// TIA Portal V20 export
// export: Created 2026-10-19T18:06:52.8062617Z, ExportSetting WithDefaults, DisplayName Totally Integrated Automation Portal, DisplayVersion V20 Update 6, DisplayName TIA Portal Openness, DisplayVersion V20 Update 6, DisplayName TIA Portal Version Control Interface, DisplayVersion V20 Update 6, DisplayName SINAMICS Startdrive Advanced, DisplayVersion V20 SP1, DisplayName SINAMICS Startdrive G130, G150, S120, S150, SINAMICS MV, G220, S200, S210, DisplayVersion V20 SP1, DisplayName SINAMICS Startdrive G110M, G120, G120C, G120D, G120P, G115D, DisplayVersion V20 SP1, DisplayName STEP 7 Professional, DisplayVersion V20 Update 6, DisplayName STEP 7 Safety, DisplayVersion V20 Update 2, DisplayName WinCC Basic/Comfort/Advanced, DisplayVersion V20 Update 6, DisplayName WinCC Unified, DisplayVersion V20 Update 6
DATA_BLOCK "SAI_IND_SpanAdjust_DB"   // DB113
VERSION : 0.1
// stored: AutoNumber true, DBAccessibleFromOPCUA true, DBAccessibleFromWebserver true, InstanceOfName SAI_IND_SpanAdjust, InstanceOfType FB
"SAI_IND_SpanAdjust"
   // VAR_INPUT
   //    ID : HW_IO;
   //    Hi_Weight : Real;
   //    Mid_Weight : Real;
   //    Low_Weight : Real;
   //    xLow_Weight : Real;
   // END_VAR
   // VAR_OUTPUT
   //    CurrentPoint : Int;
   //    CurrentWeight : Real;
   //    LoadWeight : Bool;
   //    Process : Bool;
   //    Done : Bool;
   //    Error : Bool;
   //    Cancelled : Bool;
   // END_VAR
   // VAR_IN_OUT
   //    LinearityRange : Int;
   //    Start : Bool;
   //    ConfirmWeight : Bool;
   //    Cancel : Bool;
   // END_VAR
   // VAR
   //    Activate : Bool;
   //    WRREC_SpanAdjust { S7_SetPoint := 'True'} : WRREC;
   //    RDREC_Status { S7_SetPoint := 'True'} : RDREC;
   //    IEC_Timer_1_Instance { S7_SetPoint := 'True'} : IEC_TIMER;
   //    AdjustStep : SInt;
   //    Static01 : Bool;
   //    Static02 : Bool;
   //    Static03 : Bool;
   //    Static04 : Bool;
   //    Static05 : Bool;
   //    Static06 : Bool;
   //    Static07 : Bool;
   //    Static08 : Bool;
   //    Validate_REC : SInt;
   //    Abort_REC : SInt;
   //    Check01 : Bool;
   //    Check02 : Bool;
   //    AdjustmentStatus : Int;
   //    CurrentPoint_0 : Int;
   //    CurrentWeight_0 : Real;
   // END_VAR
BEGIN
END_DATA_BLOCK
